(* IEC 61131-3 sources: avi-aoi-management/scripts/ai-eval/ngau-nhien/kho/st-tv7-canh-bao-xac-nhan/khung/src, 1 file *)

(* ---- CanhBaoXacNhan.st ---- *)
FUNCTION_BLOCK CanhBaoXacNhan
VAR_INPUT
    DIEU_KIEN : BOOL;
    XAC_NHAN : BOOL;
    T_TRE : TIME;
END_VAR
VAR_OUTPUT
    TRANG_THAI : INT;
    NHAP_NHAY : BOOL;
    CO_CANH_BAO : BOOL;
END_VAR
    (* TODO: cài đặt theo đề bài, dùng TON + R_TRIG *)
    TRANG_THAI := 0;
END_FUNCTION_BLOCK
